Staubli VAL3: resetReturnStack.pgx

public program resetReturnStack(bool x_bRecHere)
// // 清空所有记录堆栈
// // (可选)清空之后是否自动把当前点设为第一个点
  local num l_nI
  local jointRx l_jPos
  local num l_nMoveId
begin
  // ---------------------------------------------------------------------------- //
  // 清空所有记录的堆栈
  // x_bRecHere: 清空之后是否自动记录当前位置作为第一个点
  // ---------------------------------------------------------------------------- //
  //
  for l_nI= 0 to size(nMoveTypeRec)-1
    nMoveTypeRec[l_nI]=-1
    nMoveIdRec[l_nI]=-1
  endFor
  nRecIndex=0
  nCurrentMoveID=0
  bHaveGetMoveID=false

  // 是否记录当前位置为第一个点
  if x_bRecHere
    l_jPos=herej()
    call MoveJ(l_jPos,flange,mNomSpeed,l_nMoveId,false)
    waitEndMove()
  endIf

end
